(* PLC project Filler_F3, CODESYS CODESYS V3.5 SP19 3.5.19.30 *)
(* stored: creationDateTime 2024-02-20T10:41:12.000, modificationDateTime 2024-02-20T10:40:55.000 *)

PROGRAM PLC_PRG
  VAR
    Fill_Tmr : TON;  (* Fill time *)
    Start_Trig : R_TRIG;
    Running : BOOL;  (* Filler running *)
    Filling : BOOL;
  END_VAR
  VAR  (* added by the conversion: wires and edge detectors of the diagram *)
    R_TRIG1 : R_TRIG;
  END_VAR

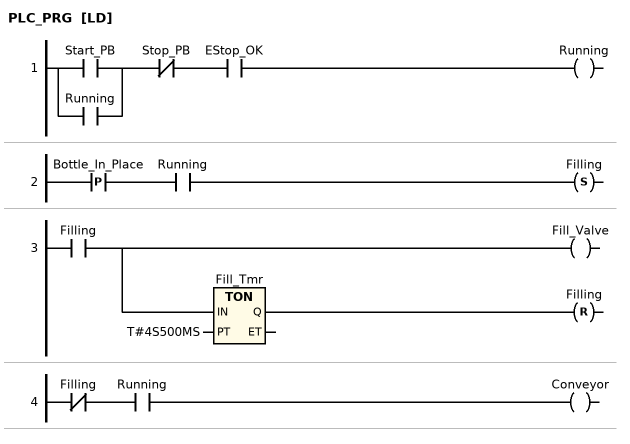
(* LD diagram, written out as Structured Text *)
Running := (Start_PB OR Running) AND NOT Stop_PB AND EStop_OK;
R_TRIG1(CLK := Bottle_In_Place);
IF R_TRIG1.Q AND Running THEN Filling := TRUE; END_IF;
Fill_Tmr(IN := Filling, PT := T#4S500MS);
Fill_Valve := Filling;
IF Fill_Tmr.Q THEN Filling := FALSE; END_IF;
Conveyor := NOT Filling AND Running;
END_PROGRAM

PROGRAM Level_Control
  VAR
    Level_Pct : REAL;  (* Bowl level, % *)
    Refill_Cnt : CTU;
  END_VAR

            (* Bowl level from the 0-10 V sensor, 0..27648 counts *)
Level_Pct := INT_TO_REAL(Level_Raw) * 100.0 / 27648.0;
IF Level_Pct < 40.0 AND Running THEN
    Refill_Valve := TRUE;
ELSIF Level_Pct > 60.0 THEN
    Refill_Valve := FALSE;
END_IF;
Refill_Cnt(CU := Refill_Valve, RESET := FALSE, PV := 1000);
FOR i := 0 TO 3 DO
    Avg[i] := 0;
END_FOR;
          
END_PROGRAM

CONFIGURATION Device
  RESOURCE Application ON PLC
    VAR_GLOBAL  (* IO_Map *)
      Start_PB AT %IX0.0 : BOOL;  (* Start push button *)
      Stop_PB AT %IX0.1 : BOOL;  (* Stop push button *)
      EStop_OK AT %IX0.2 : BOOL;  (* E-stop chain healthy *)
      Bottle_In_Place AT %IX0.3 : BOOL;  (* Bottle under the nozzle *)
      Level_Raw AT %IW2 : INT;  (* Bowl level sensor 0-10 V *)
      Fill_Valve AT %QX0.0 : BOOL;  (* Fill valve *)
      Conveyor AT %QX0.1 : BOOL;  (* Bottle conveyor *)
      Refill_Valve AT %QX0.2 : BOOL;  (* Bowl refill valve *)
    END_VAR
    TASK MainTask(INTERVAL := T#10ms, PRIORITY := 1);
    PROGRAM PLC_PRG WITH MainTask : PLC_PRG;
    PROGRAM Level_Control WITH MainTask : Level_Control;
  END_RESOURCE
END_CONFIGURATION
